(* CODESYS project Cebora.project
   CustomField04_name: CustomField04
   CustomField06_name: CustomField06
   CustomField07_name: CustomField07
   CustomField09_name: CustomField09
   CustomField08_name: CustomField08
   CustomField02_name: CustomField02
   CustomField10_name: CustomField10
   CustomField01_name: CustomField01
   CustomField03_name: CustomField03
   CustomField05_name: CustomField05

Project tree, tasks and I/O mapping:
  Cebora : TM241CEC24T/U, Schneider Electric, order no. TM241CEC24T/U, version 4.0.6.18
      settings: OPCUA enable = False
    application Application
      libraries: Toolbox, 2.2.0.0 (Schneider Electric)
      task MAST (cyclic, interval 20 ms, priority 15, watchdog 100 ms x 1) calls ConvToCAN
      global variables GVL
      program SndRecvRS232 [CFC]
      program ConvToCAN [ST]
      program Timers [LD]
    Ethernet_1 : Ethernet Network, Schneider Electric, version 4.0.6.18
    COM_Bus : COM bus, Schneider Electric, version 4.0.6.18
    Counters : Counters, Schneider Electric, version 4.0.6.18
    IO_Bus : IO bus - TM3, Schneider Electric, version 4.0.6.18
    Serial_Line_1 : Serial line, Schneider Electric, version 4.0.6.18
      ROBOT : ASCII Manager, Schneider Electric, version 4.0.0.2
    Cartridge_1 : Cartridge, Schneider Electric, version 4.0.6.18
    Pulse_Generators : Pulse Generators, Schneider Electric, version 4.0.6.18
    DQ : Digital Outputs, Schneider Electric, version 4.0.6.18
        unmapped channels: QW0, QB1
    CAN_1 : CANopen bus, Schneider Electric, version 4.0.6.18
      CANopen_Optimized : CANopen Performance, Schneider Electric, order no. 1806, version 3.0.1.24
          settings: Enable Sync generation = FALSE; Sync CobID = 126; Heartbeat in Milliseconds = 100; Enable Heartbeat generation = TRUE; Heartbeat Node ID = 100; Can Open Node ID = 100; ConfigVersion = 50659584
        CEBORA_TIG : CEBORA Power Source, CEBORA S.p.A., order no. 0, version Revision=16#00000000, FileVersion=1.2, File=CEBORA_TIG.eds
            settings: General Options.Create all SDOs = TRUE; General Options.Optional Device = TRUE; NODEIDSAVED = 3; SDO Timeout = 1000000; EXPERTSETTINGS = True; Heartbeat-Producer Time = 200; PDO 16#1400.COBID = 16#0203; PDO 16#1401.COBID = 16#0303; PDO 16#1402.COBID = 16#0403; PDO 16#1800.COBID = 16#0183; PDO 16#1800.Inhibit Time = 0; PDO 16#1800.Event Timer = 0; PDO 16#1801.COBID = 16#0283; PDO 16#1801.Inhibit Time = 0; PDO 16#1801.Event Timer = 0; PDO 16#1802.COBID = 16#0383; PDO 16#1802.Inhibit Time = 0; PDO 16#1802.Event Timer = 0; Heartbeat-Consuming1.Heartbeat-Time = 780 ms; DI0_DI7.Subindex = 16#01; DI8_DI15.Subindex = 16#02; DI16_DI23.Subindex = 16#03; DI24_D31.Subindex = 16#04; DI32_DI39.Subindex = 16#05; DI40_DI47.Subindex = 16#06; DI48_DI55.Subindex = 16#07; DI56_DI63.Subindex = 16#08; Analogue Output 1.Subindex = 16#01; Analogue Output 2.Subindex = 16#02; Analogue Output 3.Subindex = 16#03; Analogue Output 4.Subindex = 16#04; Analogue Output 5.Subindex = 16#05; Analogue Output 6.Subindex = 16#06; Analogue Output 7.Subindex = 16#07; Analogue Output 8.Subindex = 16#08; DO0_DO7.Subindex = 16#01; DO8_DO15.Subindex = 16#02; DO16_DO23.Subindex = 16#03; DO24_DO31.Subindex = 16#04; Analogue Input 1.Subindex = 16#01;
              Analogue Input 2.Subindex = 16#02; Analogue Input 3.Subindex = 16#03; Analogue Input 4.Subindex = 16#04; Analogue Input 5.Subindex = 16#05; Analogue Input 6.Subindex = 16#06; Analogue Input 7.Subindex = 16#07; Analogue Input 8.Subindex = 16#08; SDO List.Set Heartbeat Consumer.Index = 16#1016; SDO List.Set Heartbeat Consumer.Subindex = 16#01; SDO List.Set Heartbeat Consumer.Value = 16#007E030C; SDO List.Set Heartbeat Consumer.Size = 32; SDO List.Set Heartbeat Consumer.AbortIfError = FALSE; SDO List.Set Heartbeat Consumer.JumpToLine = FALSE; SDO List.Set Heartbeat Consumer.Line = 0; SDO List.Set Heartbeat Producer.Index = 16#1017; SDO List.Set Heartbeat Producer.Subindex = 16#00; SDO List.Set Heartbeat Producer.Value = 16#000000C8; SDO List.Set Heartbeat Producer.Size = 16; SDO List.Set Heartbeat Producer.AbortIfError = FALSE; SDO List.Set Heartbeat Producer.JumpToLine = FALSE; SDO List.Set Heartbeat Producer.Line = 0; SDO List.DI0_DI7.Index = 16#6200; SDO List.DI0_DI7.Subindex = 16#01; SDO List.DI0_DI7.Value = 0; SDO List.DI0_DI7.Size = 8; SDO List.DI0_DI7.AbortIfError = FALSE; SDO List.DI0_DI7.JumpToLine = FALSE; SDO List.DI0_DI7.Line = 0; SDO List.DI8_DI15.Index = 16#6200; SDO List.DI8_DI15.Subindex = 16#02; SDO List.DI8_DI15.Value = 0; SDO List.DI8_DI15.Size = 8; SDO List.DI8_DI15.AbortIfError = FALSE; SDO List.DI8_DI15.JumpToLine = FALSE; SDO List.DI8_DI15.Line = 0; SDO List.DI16_DI23.Index = 16#6200; SDO List.DI16_DI23.Subindex = 16#03; SDO List.DI16_DI23.Value = 0; SDO List.DI16_DI23.Size = 8; SDO List.DI16_DI23.AbortIfError = FALSE;
              SDO List.DI16_DI23.JumpToLine = FALSE; SDO List.DI16_DI23.Line = 0; SDO List.DI24_D31.Index = 16#6200; SDO List.DI24_D31.Subindex = 16#04; SDO List.DI24_D31.Value = 0; SDO List.DI24_D31.Size = 8; SDO List.DI24_D31.AbortIfError = FALSE; SDO List.DI24_D31.JumpToLine = FALSE; SDO List.DI24_D31.Line = 0; SDO List.DI32_DI39.Index = 16#6200; SDO List.DI32_DI39.Subindex = 16#05; SDO List.DI32_DI39.Value = 16#FF; SDO List.DI32_DI39.Size = 8; SDO List.DI32_DI39.AbortIfError = FALSE; SDO List.DI32_DI39.JumpToLine = FALSE; SDO List.DI32_DI39.Line = 0; SDO List.DI40_DI47.Index = 16#6200; SDO List.DI40_DI47.Subindex = 16#06; SDO List.DI40_DI47.Value = 0; SDO List.DI40_DI47.Size = 8; SDO List.DI40_DI47.AbortIfError = FALSE; SDO List.DI40_DI47.JumpToLine = FALSE; SDO List.DI40_DI47.Line = 0; SDO List.DI48_DI55.Index = 16#6200; SDO List.DI48_DI55.Subindex = 16#07; SDO List.DI48_DI55.Value = 0; SDO List.DI48_DI55.Size = 8; SDO List.DI48_DI55.AbortIfError = FALSE; SDO List.DI48_DI55.JumpToLine = FALSE; SDO List.DI48_DI55.Line = 0; SDO List.DI56_DI63.Index = 16#6200; SDO List.DI56_DI63.Subindex = 16#08; SDO List.DI56_DI63.Value = 0; SDO List.DI56_DI63.Size = 8; SDO List.DI56_DI63.AbortIfError = FALSE; SDO List.DI56_DI63.JumpToLine = FALSE; SDO List.DI56_DI63.Line = 0; SDO List.Analogue Output 1.Index = 16#6411; SDO List.Analogue Output 1.Subindex = 16#01; SDO List.Analogue Output 1.Value = 16#00000000;
              SDO List.Analogue Output 1.Size = 16; SDO List.Analogue Output 1.AbortIfError = FALSE; SDO List.Analogue Output 1.JumpToLine = FALSE; SDO List.Analogue Output 1.Line = 0; SDO List.Analogue Output 2.Index = 16#6411; SDO List.Analogue Output 2.Subindex = 16#02; SDO List.Analogue Output 2.Value = 16#00000000; SDO List.Analogue Output 2.Size = 16; SDO List.Analogue Output 2.AbortIfError = FALSE; SDO List.Analogue Output 2.JumpToLine = FALSE; SDO List.Analogue Output 2.Line = 0; SDO List.Analogue Output 3.Index = 16#6411; SDO List.Analogue Output 3.Subindex = 16#03; SDO List.Analogue Output 3.Value = 16#00000000; SDO List.Analogue Output 3.Size = 16; SDO List.Analogue Output 3.AbortIfError = FALSE; SDO List.Analogue Output 3.JumpToLine = FALSE; SDO List.Analogue Output 3.Line = 0; SDO List.Analogue Output 4.Index = 16#6411; SDO List.Analogue Output 4.Subindex = 16#04; SDO List.Analogue Output 4.Value = 16#00000000; SDO List.Analogue Output 4.Size = 16; SDO List.Analogue Output 4.AbortIfError = FALSE; SDO List.Analogue Output 4.JumpToLine = FALSE; SDO List.Analogue Output 4.Line = 0; SDO List.Analogue Output 5.Index = 16#6411; SDO List.Analogue Output 5.Subindex = 16#05; SDO List.Analogue Output 5.Value = 16#00000000; SDO List.Analogue Output 5.Size = 16; SDO List.Analogue Output 5.AbortIfError = FALSE; SDO List.Analogue Output 5.JumpToLine = FALSE; SDO List.Analogue Output 5.Line = 0; SDO List.Analogue Output 6.Index = 16#6411; SDO List.Analogue Output 6.Subindex = 16#06; SDO List.Analogue Output 6.Value = 16#00000000; SDO List.Analogue Output 6.Size = 16; SDO List.Analogue Output 6.AbortIfError = FALSE; SDO List.Analogue Output 6.JumpToLine = FALSE; SDO List.Analogue Output 6.Line = 0; SDO List.Analogue Output 7.Index = 16#6411;
              SDO List.Analogue Output 7.Subindex = 16#07; SDO List.Analogue Output 7.Value = 16#00000000; SDO List.Analogue Output 7.Size = 16; SDO List.Analogue Output 7.AbortIfError = FALSE; SDO List.Analogue Output 7.JumpToLine = FALSE; SDO List.Analogue Output 7.Line = 0; SDO List.Analogue Output 8.Index = 16#6411; SDO List.Analogue Output 8.Subindex = 16#08; SDO List.Analogue Output 8.Value = 16#00000000; SDO List.Analogue Output 8.Size = 16; SDO List.Analogue Output 8.AbortIfError = FALSE; SDO List.Analogue Output 8.JumpToLine = FALSE; SDO List.Analogue Output 8.Line = 0; ConfigVersion = 50659584
            output Application.CAN_SET_ArcOn : BOOL  // DI0_DI7.Bit0
            output Application.CAN_SET_RobotReady : BOOL  // DI0_DI7.Bit1
            output Application.CAN_SET_OperMode_0 : BOOL  // DI0_DI7.Bit2
            output Application.CAN_SET_OperMode_1 : BOOL  // DI0_DI7.Bit3
            output Application.CAN_SET_OperMode_2 : BOOL  // DI0_DI7.Bit4
            output Application.CAN_SET_AnalogSwap : BOOL  // DI0_DI7.Bit6
            output Application.CAN_SET_ProtocolMode : BOOL  // DI0_DI7.Bit7
            output Application.CAN_SET_GasTest : BOOL  // DI8_DI15.Bit0
            output Application.CAN_SET_WireInching : BOOL  // DI8_DI15.Bit1
            output Application.CAN_SET_WireRetract : BOOL  // DI8_DI15.Bit2
            output Application.CAN_SET_SourceErrReset : BOOL  // DI8_DI15.Bit3
            output Application.CAN_SET_TouchSensing : BOOL  // DI8_DI15.Bit4
            output Application.CAN_SET_BlowTrough : BOOL  // DI8_DI15.Bit5
            output Application.CAN_SET_JOB_0 : BOOL  // DI16_DI23.Bit0
            output Application.CAN_SET_JOB_1 : BOOL  // DI16_DI23.Bit1
            output Application.CAN_SET_JOB_2 : BOOL  // DI16_DI23.Bit2
            output Application.CAN_SET_JOB_3 : BOOL  // DI16_DI23.Bit3
            output Application.CAN_SET_JOB_4 : BOOL  // DI16_DI23.Bit4
            output Application.CAN_SET_JOB_5 : BOOL  // DI16_DI23.Bit5
            output Application.CAN_SET_JOB_6 : BOOL  // DI16_DI23.Bit6
            output Application.CAN_SET_JOB_7 : BOOL  // DI16_DI23.Bit7
            output Application.CAN_SET_WeldSim : BOOL  // DI24_D31.Bit7
            output Application.CAN_SET_AnalogSetDis_0 : BOOL  // DI32_DI39.Bit0
            output Application.CAN_SET_AnalogSetDis_1 : BOOL  // DI32_DI39.Bit1
            output Application.CAN_SET_AnalogSetDis_2 : BOOL  // DI32_DI39.Bit2
            output Application.CAN_SET_AnalogSetDis_3 : BOOL  // DI32_DI39.Bit3
            output Application.CAN_SET_AnalogSetDis_4 : BOOL  // DI32_DI39.Bit4
            output Application.CAN_SET_AnalogSetDis_5 : BOOL  // DI32_DI39.Bit5
            output Application.CAN_SET_DC_AC_Disable : BOOL  // DI40_DI47.Bit0
            output Application.CAN_SET_PLS_Disable : BOOL  // DI40_DI47.Bit3
            output Application.CAN_SET_DC_AC : BOOL  // DI48_DI55.Bit0
            output Application.CAN_SET_PLS : BOOL  // DI48_DI55.Bit3
            output Application.CAN_SET_PilotArc : BOOL  // DI48_DI55.Bit7
            output Application.CAN_SET_WeldCurrent : INT  // Analogue Output 1
            output Application.CAN_SET_WireHighSpd : INT  // Analogue Output 2
            output Application.CAN_SET_PLS_Ratio : INT  // Analogue Output 3
            output Application.CAN_SET_WireLowSpd : INT  // Analogue Output 4
            output Application.CAN_SET_PlasmaGasFlow : INT  // Analogue Output 5
            output Application.CAN_SET_ShieldGasFlow : INT  // Analogue Output 6
            input  Application.CAN_GET_CurrFlow : BOOL  // DO0_DO7.Bit0
            input  Application.CAN_GET_ProcActive : BOOL  // DO0_DO7.Bit2
            input  Application.CAN_GET_MainCurrent : BOOL  // DO0_DO7.Bit3
            input  Application.CAN_GET_CollisProtect : BOOL  // DO0_DO7.Bit4
            input  Application.CAN_GET_PowSourReady : BOOL  // DO0_DO7.Bit5
            input  Application.CAN_GET_Commun_Ready : BOOL  // DO0_DO7.Bit6
            input  Application.CAN_GET_ErrNumber_0 : BOOL  // DO8_DO15.Bit0
            input  Application.CAN_GET_ErrNumber_1 : BOOL  // DO8_DO15.Bit1
            input  Application.CAN_GET_ErrNumber_2 : BOOL  // DO8_DO15.Bit2
            input  Application.CAN_GET_ErrNumber_3 : BOOL  // DO8_DO15.Bit3
            input  Application.CAN_GET_ErrNumber_4 : BOOL  // DO8_DO15.Bit4
            input  Application.CAN_GET_ErrNumber_5 : BOOL  // DO8_DO15.Bit5
            input  Application.CAN_GET_ErrNumber_6 : BOOL  // DO8_DO15.Bit6
            input  Application.CAN_GET_ErrNumber_7 : BOOL  // DO8_DO15.Bit7
            input  Application.CAN_GET_PLS_Sync : BOOL  // DO16_DO23.Bit0
            input  Application.CAN_GET_PilotArc : BOOL  // DO16_DO23.Bit7
            input  Application.CAN_GET_StikingRem : BOOL  // DO24_DO31.Bit0
            input  Application.CAN_GET_WireAvailale : BOOL  // DO24_DO31.Bit3
            input  Application.CAN_GET_WeldVoltage : INT  // Analogue Input 1
            input  Application.CAN_GET_WeldCurrent : INT  // Analogue Input 2
            input  Application.CAN_GET_MotorCurrent : INT  // Analogue Input 3
            input  Application.CAN_GET_WireFeedSPD : INT  // Analogue Input 4
            input  Application.CAN_GET_PlasmaGasFlw : INT  // Analogue Input 5
            input  Application.CAN_GET_ShieldGasFlw : INT  // Analogue Input 6
            unmapped channels: DI0_DI7, DI8_DI15, DI16_DI23, DI24_D31, DI32_DI39, DI40_DI47, DI48_DI55, DI56_DI63, Analogue Output 7, Analogue Output 8, DO0_DO7, DO8_DO15, DO16_DO23, DO24_DO31, Analogue Input 7, Analogue Input 8
    IO : Digital Inputs, Schneider Electric, version 4.0.6.18
        unmapped channels: IW0, IB1
    Serial_Line_2 : Serial line, Schneider Electric, version 4.0.6.18
*)

// Cebora/Application/GVL
VAR_GLOBAL	
	IX0_0 AT %IX0.0:BOOL;
	InMASS:ARRAY [1..70] OF BYTE;
	InRandActual:ARRAY [1..255] OF BYTE;
	InCurrent:ARRAY [1..255] OF BYTE;
	InWireHS:ARRAY [1..255] OF BYTE;
	InPLS:ARRAY [1..255] OF BYTE;
	InWireLS:ARRAY [1..255] OF BYTE;
	InPLGAS:ARRAY [1..255] OF BYTE;
	InSHGAS:ARRAY [1..255] OF BYTE;
	InStrRandActual: STRING;
	InStrRandBefore:STRING;
	InStrCurrent:STRING;
	InStrWireHS:STRING;
	InStrPLS:STRING;
	InStrWireLS:STRING;
	InStrPLGAS:STRING;
	InStrSHGAS:STRING;
	IR_Current:REAL;
	OR_Current:REAL;
	IR_WireHS:REAL;
	OR_WireHS:REAL;
	IR_PLS:REAL;
	OR_PLS:REAL;
	IR_WireLS:REAL;
	OR_WireLS:REAL;
	IR_PLGAS:REAL;
	OR_PLGAS:REAL;
	IR_SHGAS:REAL;
	OR_SHGAS:REAL;
	I_R_PARAM:REAL;
	O_R_PARAM:REAL;	

	CAN_SET_ArcOn:BOOL;
	CAN_SET_RobotReady:BOOL;
	CAN_SET_OperMode_0:BOOL;
	CAN_SET_OperMode_1:BOOL;
	CAN_SET_OperMode_2:BOOL;
	CAN_SET_AnalogSwap:BOOL;
	CAN_SET_ProtocolMode:BOOL;
	CAN_SET_GasTest:BOOL;
	CAN_SET_WireInching:BOOL;
	CAN_SET_WireRetract:BOOL;
	CAN_SET_SourceErrReset:BOOL;
	CAN_SET_TouchSensing:BOOL;
	CAN_SET_BlowTrough:BOOL;
	CAN_SET_JOB_0:BOOL;
	CAN_SET_JOB_1:BOOL;
	CAN_SET_JOB_2:BOOL;
	CAN_SET_JOB_3:BOOL;
	CAN_SET_JOB_4:BOOL;
	CAN_SET_JOB_5:BOOL;
	CAN_SET_JOB_6:BOOL;
	CAN_SET_JOB_7:BOOL;
	CAN_SET_WeldSim:BOOL;
	CAN_SET_AnalogSetDis_0:BOOL;
	CAN_SET_AnalogSetDis_1:BOOL;
	CAN_SET_AnalogSetDis_2:BOOL;
	CAN_SET_AnalogSetDis_3:BOOL;
	CAN_SET_AnalogSetDis_4:BOOL;
	CAN_SET_AnalogSetDis_5:BOOL;
	CAN_SET_DC_AC_Disable:BOOL;
	CAN_SET_PLS_Disable:BOOL;
	CAN_SET_DC_AC:BOOL;
	CAN_SET_PLS:BOOL;
	CAN_SET_PilotArc:BOOL;
	
	CAN_SET_WeldCurrent:UINT;
	CAN_SET_WireHighSpd:UINT;
	CAN_SET_PLS_Ratio:UINT;
	CAN_SET_WireLowSpd:UINT;
	CAN_SET_PlasmaGasFlow:UINT;
	CAN_SET_ShieldGasFlow:UINT;
	
	CAN_GET_CurrFlow:BOOL;
	CAN_GET_ProcActive:BOOL;
	CAN_GET_MainCurrent:BOOL;
	CAN_GET_CollisProtect:BOOL;
	CAN_GET_PowSourReady:BOOL;
	CAN_GET_Commun_Ready:BOOL;
	CAN_GET_ErrNumber_0:BOOL;
	CAN_GET_ErrNumber_1:BOOL;
	CAN_GET_ErrNumber_2:BOOL;
	CAN_GET_ErrNumber_3:BOOL;
	CAN_GET_ErrNumber_4:BOOL;
	CAN_GET_ErrNumber_5:BOOL;
	CAN_GET_ErrNumber_6:BOOL;
	CAN_GET_ErrNumber_7:BOOL;
	CAN_GET_PLS_Sync:BOOL;
	CAN_GET_PilotArc:BOOL;
	CAN_GET_StikingRem:BOOL;
	CAN_GET_WireAvailale:BOOL;
	
	CAN_GET_WeldVoltage:UINT;
	CAN_GET_WeldCurrent:UINT;
	CAN_GET_MotorCurrent:UINT;
	CAN_GET_WireFeedSPD:UINT;
	CAN_GET_PlasmaGasFlw:UINT;
	CAN_GET_ShieldGasFlw:UINT;
	
	R_GET_WeldVoltage:REAL;
	R_GET_WeldCurrent:REAL;
	R_GET_MotorCurrent:REAL;
	R_GET_WireFeedSPD:REAL;
	R_GET_PlasmaGasFlw:REAL;
	R_GET_ShieldGasFlw:REAL;
	
	S_GET_WeldVoltage:STRING;
	S_GET_WeldCurrent:STRING;
	S_GET_MotorCurrent:STRING;
	S_GET_WireFeedSPD:STRING;
	S_GET_PlasmaGasFlw:STRING;
	S_GET_ShieldGasFlw:STRING;
	
	OutMASS:ARRAY [1..50] OF BYTE;	
	WeldVoltageMASS:ARRAY [1..255] OF BYTE;
	WeldCurrentMASS:ARRAY [1..255] OF BYTE;
	MotorCurrentMASS:ARRAY [1..255] OF BYTE;
	WireFeedSPDMASS:ARRAY [1..255] OF BYTE;
	PlasmaGasFlwMASS:ARRAY [1..255] OF BYTE;
	ShieldGasFlwMASS:ARRAY [1..255] OF BYTE;
	
	RS232Read:BOOL;
	RS232Send:BOOL;
	Readed:BOOL;
	Sended:BOOL;
	T0:TON;
	T0_STATE:BOOL;
	T1:TON;
	T1_STATE:BOOL;
	T2:TON;
	T2_STATE:BOOL;
	T3:TON;
	T3_STATE:BOOL;
	T4:TON;
	T4_ActTime:TIME;
	STOP_Read:BOOL;
	StopReadTrig:BOOL;
END_VAR

VAR_GLOBAL RETAIN
	
END_VAR

// Cebora/Application/ConvToCAN
PROGRAM ConvToCAN

VAR
	I: INT;
	FB_6: SE_TBX.FB_Scaling;
	FB_5: SE_TBX.FB_Scaling;
	FB_4: SE_TBX.FB_Scaling;
	FB_3: SE_TBX.FB_Scaling;
	FB_2: SE_TBX.FB_Scaling;
	FB_1: SE_TBX.FB_Scaling;
	FB_0: SE_TBX.FB_Scaling;;
END_VAR

IF NOT(IX0_0) THEN
	Timers();
	IF 	T0_STATE = TRUE AND Readed = FALSE THEN
		RS232Read:= TRUE;
		SndRecvRS232();
		Readed:= TRUE;
	END_IF
	Timers();
	IF T0_STATE = FALSE AND T1_STATE = TRUE THEN
		RS232Read:= FALSE;
		Readed:= FALSE;
	END_IF
	Timers();
	IF T2_STATE = TRUE AND Sended = FALSE THEN	
		RS232Send:= TRUE;
		SndRecvRS232();
		Sended:= TRUE;
	END_IF
	Timers();
	IF T1_STATE = FALSE AND T2_STATE = FALSE THEN
		RS232Send:= FALSE;
		Sended:= FALSE;
	END_IF
	
	FOR I:= 1 TO 5 BY 1 DO
		InRandActual[I]:= InMASS[I+64];
	END_FOR
	
	InStrRandActual:= ArrayOfByte_TO_String(i_abyIput:= InRandActual, i_xOrdr:= TRUE , i_xSpce:=  FALSE);
	IF 	InStrRandActual = InStrRandBefore THEN
		StopReadTrig:= TRUE;
	ELSE
		StopReadTrig:= FALSE;
	END_IF
	
	//Reading data
	IF 	STOP_Read = TRUE THEN
		FOR I:= 1 TO 70 BY 1 DO
			InMASS[I]:= 48;
		END_FOR
	END_IF
	
	IF 	InMASS[1] = 83 AND InMASS[70] = 70 OR STOP_Read = TRUE THEN
		IF 	InMASS[2] = 49 THEN
			CAN_SET_ArcOn:= TRUE;
		ELSE
			CAN_SET_ArcOn:= FALSE;
		END_IF
		IF 	InMASS[3] = 49 THEN
			CAN_SET_RobotReady:= TRUE;
		ELSE
			CAN_SET_RobotReady:= FALSE;
		END_IF
		IF 	InMASS[4] = 49 THEN
			CAN_SET_OperMode_0:= TRUE;
		ELSE
			CAN_SET_OperMode_0:= FALSE;
		END_IF
		IF 	InMASS[5] = 49 THEN
			CAN_SET_OperMode_1:= TRUE;
		ELSE
			CAN_SET_OperMode_1:= FALSE;
		END_IF
		IF 	InMASS[6] = 49 THEN
			CAN_SET_OperMode_2:= TRUE;
		ELSE
			CAN_SET_OperMode_2:= FALSE;
		END_IF
		IF 	InMASS[7] = 49 THEN
			CAN_SET_AnalogSwap:= TRUE;
		ELSE
			CAN_SET_AnalogSwap:= FALSE;
		END_IF
		IF 	InMASS[8] = 49 THEN
			CAN_SET_ProtocolMode:= TRUE;
		ELSE
			CAN_SET_ProtocolMode:= FALSE;
		END_IF
		IF 	InMASS[9] = 49 THEN
			CAN_SET_GasTest:= TRUE;
		ELSE
			CAN_SET_GasTest:= FALSE;
		END_IF
		IF 	InMASS[10] = 49 THEN
			CAN_SET_WireInching:= TRUE;
		ELSE
			CAN_SET_WireInching:= FALSE;
		END_IF
		IF 	InMASS[11] = 49 THEN
			CAN_SET_WireRetract:= TRUE;
		ELSE
			CAN_SET_WireRetract:= FALSE;
		END_IF
		IF 	InMASS[12] = 49 THEN
			CAN_SET_SourceErrReset:= TRUE;
		ELSE
			CAN_SET_SourceErrReset:= FALSE;
		END_IF
		IF 	InMASS[13] = 49 THEN
			CAN_SET_TouchSensing:= TRUE;
		ELSE
			CAN_SET_TouchSensing:= FALSE;
		END_IF
		IF 	InMASS[14] = 49 THEN
			CAN_SET_BlowTrough:= TRUE;
		ELSE
			CAN_SET_BlowTrough:= FALSE;
		END_IF
		IF 	InMASS[15] = 49 THEN
			CAN_SET_JOB_0:= TRUE;
		ELSE
			CAN_SET_JOB_0:= FALSE;
		END_IF
		IF 	InMASS[16] = 49 THEN
			CAN_SET_JOB_1:= TRUE;
		ELSE
			CAN_SET_JOB_1:= FALSE;
		END_IF
		IF 	InMASS[17] = 49 THEN
			CAN_SET_JOB_2:= TRUE;
		ELSE
			CAN_SET_JOB_2:= FALSE;
		END_IF
		IF 	InMASS[18] = 49 THEN
			CAN_SET_JOB_3:= TRUE;
		ELSE
			CAN_SET_JOB_3:= FALSE;
		END_IF
		IF 	InMASS[19] = 49 THEN
			CAN_SET_JOB_4:= TRUE;
		ELSE
			CAN_SET_JOB_4:= FALSE;
		END_IF
		IF 	InMASS[20] = 49 THEN
			CAN_SET_JOB_5:= TRUE;
		ELSE
			CAN_SET_JOB_5:= FALSE;
		END_IF
		IF 	InMASS[21] = 49 THEN
			CAN_SET_JOB_6:= TRUE;
		ELSE
			CAN_SET_JOB_6:= FALSE;
		END_IF
		IF 	InMASS[22] = 49 THEN
			CAN_SET_JOB_7:= TRUE;
		ELSE
			CAN_SET_JOB_7:= FALSE;
		END_IF
		IF 	InMASS[23] = 49 THEN
			CAN_SET_WeldSim:= TRUE;
		ELSE
			CAN_SET_WeldSim:= FALSE;
		END_IF
		IF 	InMASS[24] = 49 THEN
			CAN_SET_AnalogSetDis_0:= TRUE;
		ELSE
			CAN_SET_AnalogSetDis_0:= FALSE;
		END_IF
		IF 	InMASS[25] = 49 THEN
			CAN_SET_AnalogSetDis_1:= TRUE;
		ELSE
			CAN_SET_AnalogSetDis_1:= FALSE;
		END_IF
		IF 	InMASS[26] = 49 THEN
			CAN_SET_AnalogSetDis_2:= TRUE;
		ELSE
			CAN_SET_AnalogSetDis_2:= FALSE;
		END_IF
		IF 	InMASS[27] = 49 THEN
			CAN_SET_AnalogSetDis_3:= TRUE;
		ELSE
			CAN_SET_AnalogSetDis_3:= FALSE;
		END_IF
		IF 	InMASS[28] = 49 THEN
			CAN_SET_AnalogSetDis_4:= TRUE;
		ELSE
			CAN_SET_AnalogSetDis_4:= FALSE;
		END_IF
		IF 	InMASS[29] = 49 THEN
			CAN_SET_AnalogSetDis_5:= TRUE;
		ELSE
			CAN_SET_AnalogSetDis_5:= FALSE;
		END_IF
		IF 	InMASS[30] = 49 THEN
			CAN_SET_DC_AC_Disable:= TRUE;
		ELSE
			CAN_SET_DC_AC_Disable:= FALSE;
		END_IF
		IF 	InMASS[31] = 49 THEN
			CAN_SET_PLS_Disable:= TRUE;
		ELSE
			CAN_SET_PLS_Disable:= FALSE;
		END_IF
		IF 	InMASS[32] = 49 THEN
			CAN_SET_DC_AC:= TRUE;
		ELSE
			CAN_SET_DC_AC:= FALSE;
		END_IF
		IF 	InMASS[33] = 49 THEN
			CAN_SET_PLS:= TRUE;
		ELSE
			CAN_SET_PLS:= FALSE;
		END_IF
		IF 	InMASS[34] = 49 THEN
			CAN_SET_PilotArc:= TRUE;
		ELSE
			CAN_SET_PilotArc:= FALSE;
		END_IF
		FOR I:= 1 TO 5 BY 1 DO
			InCurrent[I]:= InMASS[I+34];
			InWireHS[I]:= InMASS[I+39];
			InPLS[I]:= InMASS[I+44];
			InWireLS[I]:= InMASS[I+49];
			InPLGAS[I]:= InMASS[I+54];
			InSHGAS[I]:= InMASS[I+59];
		END_FOR
		InStrCurrent:= ArrayOfByte_TO_String(i_abyIput:= InCurrent, i_xOrdr:= TRUE , i_xSpce:=  FALSE);
		InStrWireHS:= ArrayOfByte_TO_String(i_abyIput:= InWireHS, i_xOrdr:= TRUE , i_xSpce:=  FALSE);
		InStrPLS:= ArrayOfByte_TO_String(i_abyIput:= InPLS, i_xOrdr:= TRUE , i_xSpce:=  FALSE);
		InStrWireLS:= ArrayOfByte_TO_String(i_abyIput:= InWireLS, i_xOrdr:= TRUE , i_xSpce:=  FALSE);
		InStrPLGAS:= ArrayOfByte_TO_String(i_abyIput:= InPLGAS, i_xOrdr:= TRUE , i_xSpce:=  FALSE);
		InStrSHGAS:= ArrayOfByte_TO_String(i_abyIput:= InSHGAS, i_xOrdr:= TRUE , i_xSpce:=  FALSE);
		//Set Current
		IR_Current:= STRING_TO_REAL(InStrCurrent);
		FB_0( i_xEn:= TRUE,i_rIput:= IR_Current,i_rMinIput:= 0.0,i_rMaxIput:= 500.0,i_rMinOput:= 0.0,i_rMaxOput:= 65535.0,q_rOput=> OR_Current);
		CAN_SET_WeldCurrent:= REAL_TO_UINT(OR_Current);
		//Set Wire High Speed
		IR_WireHS:= STRING_TO_REAL(InStrWireHS);
		FB_0( i_xEn:= TRUE,i_rIput:= IR_WireHS,i_rMinIput:= -10.0,i_rMaxIput:= 10.0,i_rMinOput:= 0.0,i_rMaxOput:= 65535.0,q_rOput=> OR_WireHS);
		CAN_SET_WireHighSpd:= REAL_TO_UINT(OR_WireHS);
		//Set Pulse Raito
		IR_PLS:= STRING_TO_REAL(InStrPLS);
		FB_0( i_xEn:= TRUE,i_rIput:= IR_PLS,i_rMinIput:= 0.0,i_rMaxIput:= 100.0,i_rMinOput:= 0.0,i_rMaxOput:= 65535.0,q_rOput=> OR_PLS);
		CAN_SET_PLS_Ratio:= REAL_TO_UINT(OR_PLS);
		//Set Wire Low Speed
		IR_WireLS:= STRING_TO_REAL(InStrWireLS);
		FB_0( i_xEn:= TRUE,i_rIput:= IR_WireLS,i_rMinIput:= -10.0,i_rMaxIput:= 10.0,i_rMinOput:= 0.0,i_rMaxOput:= 65535.0,q_rOput=> OR_WireLS);
		CAN_SET_WireLowSpd:= REAL_TO_UINT(OR_WireLS);	
		//Set Plasma Gas Flow
		IR_PLGAS:= STRING_TO_REAL(InStrPLGAS);
		FB_0( i_xEn:= TRUE,i_rIput:= IR_PLGAS,i_rMinIput:= 0.0,i_rMaxIput:= 10.0,i_rMinOput:= 0.0,i_rMaxOput:= 65535.0,q_rOput=> OR_PLGAS);
		CAN_SET_PlasmaGasFlow:= REAL_TO_UINT(OR_PLGAS);	
		//Set Shield Gas Flow
		IR_SHGAS:= STRING_TO_REAL(InStrSHGAS);
		FB_0( i_xEn:= TRUE,i_rIput:= IR_SHGAS,i_rMinIput:= 0.0,i_rMaxIput:= 30.0,i_rMinOput:= 0.0,i_rMaxOput:= 65535.0,q_rOput=> OR_SHGAS);
		CAN_SET_ShieldGasFlow:= REAL_TO_UINT(OR_SHGAS);
	END_IF
	//Reading data
	
	//Sending data
	OutMASS[1]:= 83;
	IF 	CAN_GET_CurrFlow = TRUE THEN
		OutMASS[2]:= 49;
	ELSE
		OutMASS[2]:= 48;
	END_IF
	IF 	CAN_GET_ProcActive = TRUE THEN
		OutMASS[3]:= 49;
	ELSE
		OutMASS[3]:= 48;
	END_IF
	IF 	CAN_GET_MainCurrent = TRUE THEN
		OutMASS[4]:= 49;
	ELSE
		OutMASS[4]:= 48;
	END_IF
	IF 	CAN_GET_CollisProtect = TRUE THEN
		OutMASS[5]:= 49;
	ELSE
		OutMASS[5]:= 48;
	END_IF
	IF 	CAN_GET_PowSourReady = TRUE THEN
		OutMASS[6]:= 49;
	ELSE
		OutMASS[6]:= 48;
	END_IF
	IF 	CAN_GET_Commun_Ready = TRUE THEN
		OutMASS[7]:= 49;
	ELSE
		OutMASS[7]:= 48;
	END_IF
	IF 	CAN_GET_ErrNumber_0 = TRUE THEN
		OutMASS[8]:= 49;
	ELSE
		OutMASS[8]:= 48;
	END_IF
	IF 	CAN_GET_ErrNumber_1 = TRUE THEN
		OutMASS[9]:= 49;
	ELSE
		OutMASS[9]:= 48;
	END_IF
	IF 	CAN_GET_ErrNumber_2 = TRUE THEN
		OutMASS[10]:= 49;
	ELSE
		OutMASS[10]:= 48;
	END_IF
	IF 	CAN_GET_ErrNumber_3 = TRUE THEN
		OutMASS[11]:= 49;
	ELSE
		OutMASS[11]:= 48;
	END_IF
	IF 	CAN_GET_ErrNumber_4 = TRUE THEN
		OutMASS[12]:= 49;
	ELSE
		OutMASS[12]:= 48;
	END_IF
	IF 	CAN_GET_ErrNumber_5 = TRUE THEN
		OutMASS[13]:= 49;
	ELSE
		OutMASS[13]:= 48;
	END_IF
	IF 	CAN_GET_ErrNumber_6 = TRUE THEN
		OutMASS[14]:= 49;
	ELSE
		OutMASS[14]:= 48;
	END_IF
	IF 	CAN_GET_ErrNumber_7 = TRUE THEN
		OutMASS[15]:= 49;
	ELSE
		OutMASS[15]:= 48;
	END_IF
	IF 	CAN_GET_PLS_Sync = TRUE THEN
		OutMASS[16]:= 49;
	ELSE
		OutMASS[16]:= 48;
	END_IF
	IF 	CAN_GET_PilotArc = TRUE THEN
		OutMASS[17]:= 49;
	ELSE
		OutMASS[17]:= 48;
	END_IF
	IF 	CAN_GET_StikingRem = TRUE THEN
		OutMASS[18]:= 49;
	ELSE
		OutMASS[18]:= 48;
	END_IF
	IF 	CAN_GET_WireAvailale = TRUE THEN
		OutMASS[19]:= 49;
	ELSE
		OutMASS[19]:= 48;
	END_IF
	
	FB_1( i_xEn:= TRUE,i_rIput:= UINT_TO_REAL(CAN_GET_WeldVoltage),i_rMinIput:= 0.0,i_rMaxIput:= 65535.0,i_rMinOput:= 0.0,i_rMaxOput:= 100.0,q_rOput=> R_GET_WeldVoltage);
	FB_2( i_xEn:= TRUE,i_rIput:= UINT_TO_REAL(CAN_GET_WeldCurrent),i_rMinIput:= 0.0,i_rMaxIput:= 65535.0,i_rMinOput:= 0.0,i_rMaxOput:= 1000.0,q_rOput=> R_GET_WeldCurrent);
	FB_3( i_xEn:= TRUE,i_rIput:= UINT_TO_REAL(CAN_GET_MotorCurrent),i_rMinIput:= 0.0,i_rMaxIput:= 65535.0,i_rMinOput:= 0.0,i_rMaxOput:= 5.0,q_rOput=> R_GET_MotorCurrent);
	FB_4( i_xEn:= TRUE,i_rIput:= UINT_TO_REAL(CAN_GET_WireFeedSPD),i_rMinIput:= 0.0,i_rMaxIput:= 65535.0,i_rMinOput:= -12.5,i_rMaxOput:= 12.5,q_rOput=> R_GET_WireFeedSPD);
	FB_5( i_xEn:= TRUE,i_rIput:= UINT_TO_REAL(CAN_GET_PlasmaGasFlw),i_rMinIput:= 0.0,i_rMaxIput:= 65535.0,i_rMinOput:= 0.0,i_rMaxOput:= 10.0,q_rOput=> R_GET_PlasmaGasFlw);
	FB_6( i_xEn:= TRUE,i_rIput:= UINT_TO_REAL(CAN_GET_ShieldGasFlw),i_rMinIput:= 0.0,i_rMaxIput:= 65535.0,i_rMinOput:= 0.0,i_rMaxOput:= 30.0,q_rOput=> R_GET_ShieldGasFlw);
	S_GET_WeldVoltage:= REAL_TO_STRING(R_GET_WeldVoltage);
	S_GET_WeldCurrent:= REAL_TO_STRING(R_GET_WeldCurrent);
	S_GET_MotorCurrent:= REAL_TO_STRING(R_GET_MotorCurrent);
	S_GET_WireFeedSPD:= REAL_TO_STRING(R_GET_WireFeedSPD);
	S_GET_PlasmaGasFlw:= REAL_TO_STRING(R_GET_PlasmaGasFlw);
	S_GET_ShieldGasFlw:= REAL_TO_STRING(R_GET_ShieldGasFlw);
	WeldVoltageMASS:= String_TO_ArrayOfByte(i_sIput:= S_GET_WeldVoltage,i_xOrdr:= TRUE);
	WeldCurrentMASS:= String_TO_ArrayOfByte(i_sIput:= S_GET_WeldCurrent,i_xOrdr:= TRUE);
	MotorCurrentMASS:= String_TO_ArrayOfByte(i_sIput:= S_GET_MotorCurrent,i_xOrdr:= TRUE);
	WireFeedSPDMASS:= String_TO_ArrayOfByte(i_sIput:= S_GET_WireFeedSPD,i_xOrdr:= TRUE);
	PlasmaGasFlwMASS:= String_TO_ArrayOfByte(i_sIput:= S_GET_PlasmaGasFlw,i_xOrdr:= TRUE);
	ShieldGasFlwMASS:= String_TO_ArrayOfByte(i_sIput:= S_GET_ShieldGasFlw,i_xOrdr:= TRUE);
	
	FOR I:= 1 TO 5 BY 1 DO
		OutMASS[I+19]:= WeldVoltageMASS[I];
		OutMASS[I+24]:= WeldCurrentMASS[I];
		OutMASS[I+29]:= MotorCurrentMASS[I];
		OutMASS[I+34]:= WireFeedSPDMASS[I];
		OutMASS[I+39]:= PlasmaGasFlwMASS[I];
		OutMASS[I+44]:= ShieldGasFlwMASS[I];
	END_FOR;
	
	IF 	LEN(S_GET_WeldVoltage) = 3 THEN
		OutMASS[23]:= 48;
		OutMASS[24]:= 48;
	ELSIF LEN(S_GET_WeldVoltage) = 4 THEN
		OutMASS[24]:= 48;
	END_IF
	IF 	LEN(S_GET_WeldCurrent) = 3 THEN
		OutMASS[28]:= 48;
		OutMASS[29]:= 48;
	ELSIF LEN(S_GET_WeldCurrent) = 4 THEN
		OutMASS[29]:= 48;
	END_IF
	IF 	LEN(S_GET_MotorCurrent) = 3 THEN
		OutMASS[33]:= 48;
		OutMASS[34]:= 48;
	ELSIF LEN(S_GET_MotorCurrent) = 4 THEN
		OutMASS[34]:= 48;
	END_IF
	IF 	LEN(S_GET_WireFeedSPD) = 3 THEN
		OutMASS[38]:= 48;
		OutMASS[39]:= 48;
	ELSIF LEN(S_GET_WireFeedSPD) = 4 THEN
		OutMASS[39]:= 48;
	END_IF
	IF 	LEN(S_GET_PlasmaGasFlw) = 3 THEN
		OutMASS[43]:= 48;
		OutMASS[44]:= 48;
	ELSIF LEN(S_GET_PlasmaGasFlw) = 4 THEN
		OutMASS[44]:= 48;
	END_IF
	IF 	LEN(S_GET_ShieldGasFlw) = 3 THEN
		OutMASS[48]:= 48;
		OutMASS[49]:= 48;
	ELSIF LEN(S_GET_ShieldGasFlw) = 4 THEN
		OutMASS[49]:= 48;
	END_IF
	OutMASS[50]:= 70;
	//Sending data
	InStrRandBefore:= InStrRandActual;
END_IF

END_PROGRAM

// Cebora/Application/Timers
PROGRAM Timers
VAR
END_VAR

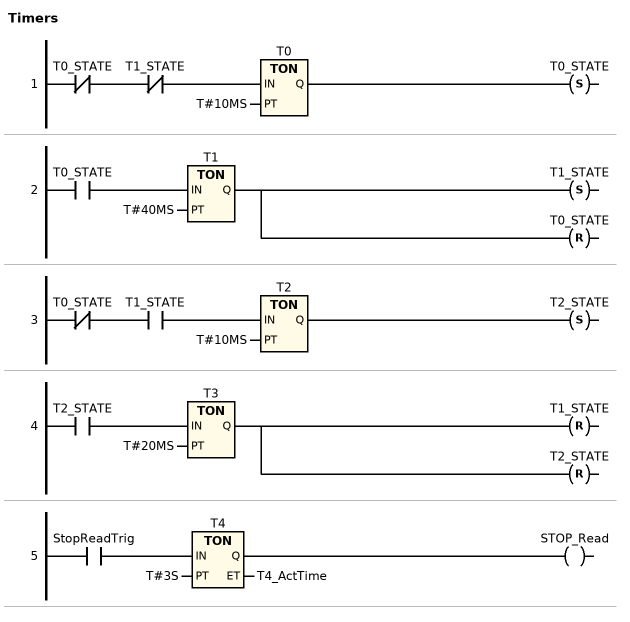
// NETWORK 1
T0(IN := NOT T0_STATE AND NOT T1_STATE, PT := T#10MS); // TON
T0_STATE S= T0.Q;

// NETWORK 2
T1(IN := T0_STATE, PT := T#40MS); // TON
T1_STATE S= T1.Q;
T0_STATE R= T1.Q;

// NETWORK 3
T2(IN := NOT T0_STATE AND T1_STATE, PT := T#10MS); // TON
T2_STATE S= T2.Q;

// NETWORK 4
T3(IN := T2_STATE, PT := T#20MS); // TON
T1_STATE R= T3.Q;
T2_STATE R= T3.Q;

// NETWORK 5
T4(IN := StopReadTrig, PT := T#3S, ET => T4_ActTime); // TON
STOP_Read := T4.Q;

END_PROGRAM

// Cebora/Application/SndRecvRS232
PROGRAM SndRecvRS232
VAR
	ADDM1: ADDM;
	ADDM2: ADDM;
	myAddressTable: ADDRESS;
	RS232_READ: SEND_RECV_MSG;
	RS232_SEND: SEND_RECV_MSG;
END_VAR

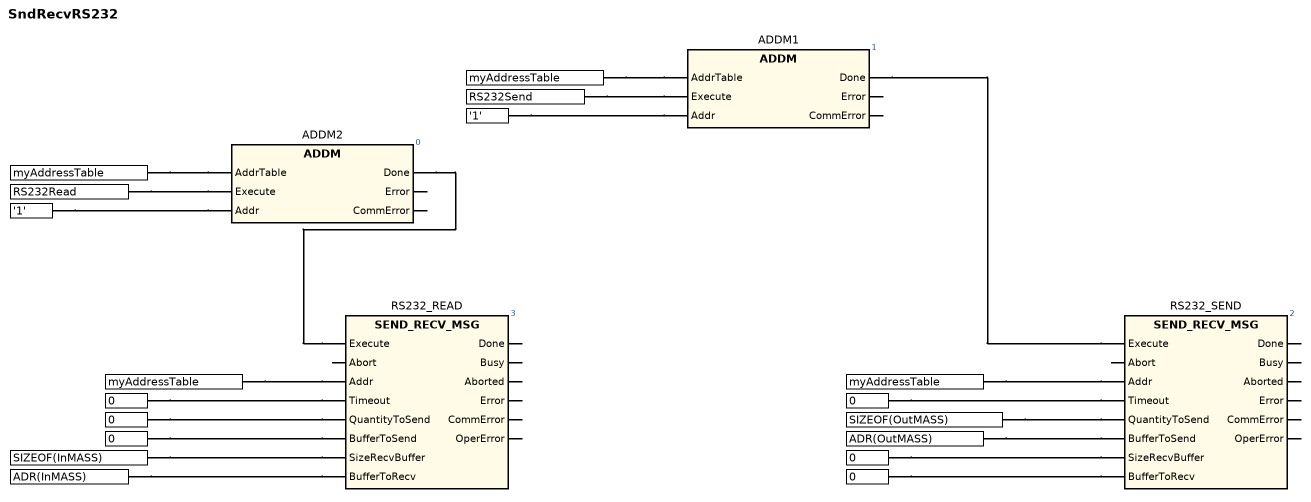
ADDM2(AddrTable := myAddressTable, Execute := RS232Read, Addr := '1'); // ADDM
ADDM1(AddrTable := myAddressTable, Execute := RS232Send, Addr := '1'); // ADDM
RS232_SEND(
    Execute := ADDM1.Done,
    Addr := myAddressTable,
    Timeout := 0,
    QuantityToSend := SIZEOF(OutMASS),
    BufferToSend := ADR(OutMASS),
    SizeRecvBuffer := 0,
    BufferToRecv := 0); // SEND_RECV_MSG
RS232_READ(
    Execute := ADDM2.Done,
    Addr := myAddressTable,
    Timeout := 0,
    QuantityToSend := 0,
    BufferToSend := 0,
    SizeRecvBuffer := SIZEOF(InMASS),
    BufferToRecv := ADR(InMASS)); // SEND_RECV_MSG

END_PROGRAM
